(* IEC 61131-3 sources: plc-hackathon-2026/work/dump/MyController/Plc Logic/Application/CustomTypes, 6 files *)

(* ---- typeAgg.st ---- *)
TYPE typeAgg:
// VERSION : 0.1
// ---------------------------------------------------------------------
// Agregirane energije [kWh] i troskovi [EUR] - LReal zbog preciznosti
// ---------------------------------------------------------------------
   STRUCT
      E_fne : LReal;   // ostvarena proizvodnja FNE (nakon curtailmenta)
      E_fne_curtailed : LReal;   // energija odrezana curtailmentom
      E_fec : LReal;   // fiksna potrosnja
      E_bess_chg : LReal;   // punjenje baterije (sa strane sabirnice)
      E_bess_dch : LReal;   // praznjenje baterije (sa strane sabirnice)
      E_ev : LReal;   // energija na sabirnici predana punjacima
      E_ev_required : LReal;   // zatrazena energija (sesije zapoceta u periodu)
      E_ev_unmet : LReal;   // nepredana energija pri odlasku vozila
      E_import : LReal;
      E_export : LReal;
      P_peak : LReal;   // max snaga uvoza na 15-min intervalu [kW]
      cost_energy : LReal;   // trosak energije (uvoz - izvoz)
      cost_grid : LReal;   // mrezarina
      cost_peak : LReal;   // trosak vrsne snage
      cost_total : LReal;
   END_STRUCT
END_TYPE

(* ---- typeEVCmd.st ---- *)
TYPE typeEVCmd:
// VERSION : 0.1
// ---------------------------------------------------------------------
// Sucelje: ulazi simulatora (pise regulator)
// ---------------------------------------------------------------------
   STRUCT
      P_charge : Real;   // [kW]
   END_STRUCT
END_TYPE

(* ---- typeEVOut.st ---- *)
TYPE typeEVOut:
// VERSION : 0.1
// ---------------------------------------------------------------------
// Sucelje: izlazi simulatora (cita regulator)
// ---------------------------------------------------------------------
   STRUCT
      connected : Bool;
      planned_departure : DT;   // (odlazak iza kraja godine je ogranicen na zadnji korak)
      PD_DT_YEAR : UINT;
	  PD_DT_MONTH : USINT;
	  PD_DT_DAY : USINT;
	  PD_DT_WEEKDAY : USINT;
	  PD_DT_HOUR : USINT;
	  PD_DT_MINUTE : USINT;
	  PD_DT_SECOND : USINT;
	  PD_DT_NANOSECOND : USINT;
	  energy_required : REAL;   // [kWh] jos treba dostaviti (E* - E)
      energy_delivered : Real;   // [kWh] dostavljeno u sesiji
      P_charge_act : Real;   // [kW] ostvarena snaga u PROSLOM koraku
   END_STRUCT
END_TYPE

(* ---- typeSimCmd.st ---- *)
TYPE typeSimCmd:
// VERSION : 0.1
   STRUCT
      FNE_enable_curtail : BOOL;
      FNE_curtail_value : REAL;   // [kW]
      BESS_enable_charge : BOOL;
      BESS_P_charge : REAL;   // [kW]
      BESS_enable_discharge : BOOL;
      BESS_P_discharge : REAL;   // [kW]
      EV : Array[0..3] of typeEVCmd;
   END_STRUCT
END_TYPE

(* ---- typeSimOut.st ---- *)
TYPE typeSimOut:
// VERSION : 0.1
   STRUCT
      t_sim : typeSimTime;
      FNE_output_power : Real;   // [kW] RASPOLOZIVA snaga u intervalu k (prije curtailmenta)
      FNE_P_act : Real;   // [kW] ostvarena snaga u proslom koraku
      FEC_P_fix : Real;   // [kW] fiksna potrosnja u intervalu k
      BESS_SoC : Real;   // [%] na pocetku intervala k
      BESS_P_charge_act : Real;   // [kW] ostvareno u proslom koraku
      BESS_P_discharge_act : Real;   // [kW] ostvareno u proslom koraku
      EV : ARRAY[0..3] OF typeEVOut;
      EGC_P_import : Real;   // [kW] izmjereno u PROSLOM koraku (k-1)
      EGC_P_export : Real;   // [kW] izmjereno u PROSLOM koraku (k-1)
      EGC_overload_import : Bool;
      EGC_overload_export : Bool;
      sim_finished : Bool;
      sim_tripped : Bool;   // postrojenje odspojeno (overload) - latch
   END_STRUCT
END_TYPE

(* ---- typeSimTime.st ---- *)
TYPE typeSimTime:
// ---------------------------------------------------------------------
// Simulirano vrijeme (izvedeno iz brojaca koraka k)
// ---------------------------------------------------------------------
	STRUCT
		k : DINT;   // indeks koraka 0..35039
		DT_YEAR : UINT;
		DT_MONTH : USINT;
		DT_DAY : USINT;
		DT_WEEKDAY : USINT;
		DT_HOUR : USINT;
		DT_MINUTE : USINT;
		DT_SECOND : USINT;
		DT_NANOSECOND : USINT;
		stamp : DT;   // simulirani datum/vrijeme POCETKA intervala
		qh_of_day : Int;   // 0..95
		day_of_year : Int;   // 0..364
		month : Int;   // 1..12
		weekday : Int;   // 1=pon .. 7=ned
		tariff_high : Bool;   // TRUE = visa tarifa (VT)
	END_STRUCT
END_TYPE
